Fanuc KAREL source: KT00793.KL

PROGRAM KT00793
%NOLOCKGROUP
VAR
  B1: BOOLEAN
  B2: BOOLEAN
  OUT: REAL
BEGIN
  B1 = TRUE
  B2 = FALSE
  B1 = TRUE
  B2 = FALSE
  OUT = COS(B1)
END KT00793
